Fanuc KAREL source: kb00122.KL

-- PROVISIONAL review KL for V1013-1; original PC SHA256 f3ac6aa9c2f6016a5f83166252d13d3410a5ab9f824302e72932369e734603d6
-- Incomplete behavior may be omitted. Consult companion uncertainty JSON. Do not deploy.
PROGRAM KB00122
%NOLOCKGROUP
BEGIN
  -- UNRESOLVED_PC offsets 5-14; opcodes 3F,75
  -- UNRESOLVED_PC offsets 19-26; opcodes 9D,23
  -- UNRESOLVED_PC offsets 31-49; opcodes 27,22,2A,22,31
  -- UNRESOLVED_PC offsets 54-58; opcodes 7F
END KB00122
